// TIA Portal V17 program export: 1 tag tables, 0 data types, 1 data blocks, 1 code blocks (in call order from the OBs), 0 instance data blocks

VAR_GLOBAL   // PLC tag table "红绿灯变量表"
   StartPB AT %M0.0 : Bool;   // HMI 启动按钮
   StopPB AT %M0.1 : Bool;   // HMI 停止按钮
   Run AT %M0.2 : Bool;   // 运行自锁与指示灯
   NS_Red AT %Q0.0 : Bool;   // 南北红灯
   NS_Yellow AT %Q0.1 : Bool;   // 南北黄灯
   NS_Green AT %Q0.2 : Bool;   // 南北绿灯
   EW_Red AT %Q0.3 : Bool;   // 东西红灯
   EW_Yellow AT %Q0.4 : Bool;   // 东西黄灯
   EW_Green AT %Q0.5 : Bool;   // 东西绿灯
   Done1 AT %M1.0 : Bool;   // 东西绿灯定时到
   Done2 AT %M1.1 : Bool;   // 东西黄灯定时到
   Done3 AT %M1.2 : Bool;   // 南北绿灯定时到
   Done4 AT %M1.3 : Bool;   // 南北黄灯定时到
END_VAR

DATA_BLOCK "TrafficTimers"   // DB1
{ S7_Optimized_Access := 'FALSE' }
   VAR
      T1 : TON_TIME;
      T2 : TON_TIME;
      T3 : TON_TIME;
      T4 : TON_TIME;
   END_VAR
BEGIN
END_DATA_BLOCK

ORGANIZATION_BLOCK "Main"   // OB1, LAD, ProgramCycle
{ S7_Optimized_Access := 'TRUE' }
VERSION : 0.1
// stored: AutoNumber true, IsIECCheckEnabled false, SetENOAutomatically false
   VAR_INPUT
      Initial_Call : Bool;   // Initial call of this OB
      Remanence : Bool;   // =True, if remanent data are available
   END_VAR
BEGIN

REGION Network 1: 启停自锁
   // 启动后保持运行，停止优先。
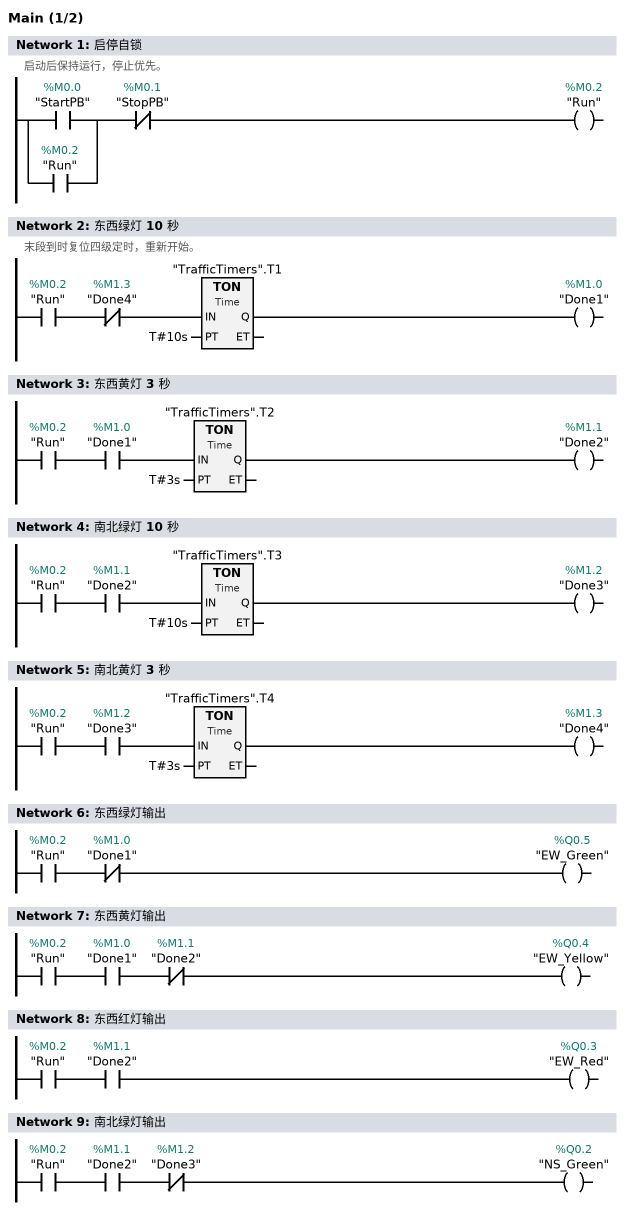
   RUNG wire#powerrail
      Contact( "StartPB" )
      wire#w1
      I_Contact( "StopPB" )
      Coil( "Run" )
   END_RUNG
   RUNG wire#powerrail
      Contact( "Run" )
   END_RUNG wire#w1
   // the same network as SCL:
   "Run" := ("StartPB" OR "Run") AND NOT "StopPB";
END_REGION

REGION Network 2: 东西绿灯 10 秒
   // 末段到时复位四级定时，重新开始。
   RUNG wire#powerrail
      Contact( "Run" )
      I_Contact( "Done4" )
      { S7_Templates := "time_type := Time" } "TrafficTimers".T1.TON(pt := T#10s, et =>)
      Coil( "Done1" )
   END_RUNG
   // the same network as SCL:
   "TrafficTimers".T1.TON(IN := "Run" AND NOT "Done4", PT := T#10s);
   "Done1" := "TrafficTimers".T1.Q;
END_REGION

REGION Network 3: 东西黄灯 3 秒
   RUNG wire#powerrail
      Contact( "Run" )
      Contact( "Done1" )
      { S7_Templates := "time_type := Time" } "TrafficTimers".T2.TON(pt := T#3s, et =>)
      Coil( "Done2" )
   END_RUNG
   // the same network as SCL:
   "TrafficTimers".T2.TON(IN := "Run" AND "Done1", PT := T#3s);
   "Done2" := "TrafficTimers".T2.Q;
END_REGION

REGION Network 4: 南北绿灯 10 秒
   RUNG wire#powerrail
      Contact( "Run" )
      Contact( "Done2" )
      { S7_Templates := "time_type := Time" } "TrafficTimers".T3.TON(pt := T#10s, et =>)
      Coil( "Done3" )
   END_RUNG
   // the same network as SCL:
   "TrafficTimers".T3.TON(IN := "Run" AND "Done2", PT := T#10s);
   "Done3" := "TrafficTimers".T3.Q;
END_REGION

REGION Network 5: 南北黄灯 3 秒
   RUNG wire#powerrail
      Contact( "Run" )
      Contact( "Done3" )
      { S7_Templates := "time_type := Time" } "TrafficTimers".T4.TON(pt := T#3s, et =>)
      Coil( "Done4" )
   END_RUNG
   // the same network as SCL:
   "TrafficTimers".T4.TON(IN := "Run" AND "Done3", PT := T#3s);
   "Done4" := "TrafficTimers".T4.Q;
END_REGION

REGION Network 6: 东西绿灯输出
   RUNG wire#powerrail
      Contact( "Run" )
      I_Contact( "Done1" )
      Coil( "EW_Green" )
   END_RUNG
   // the same network as SCL:
   "EW_Green" := "Run" AND NOT "Done1";
END_REGION

REGION Network 7: 东西黄灯输出
   RUNG wire#powerrail
      Contact( "Run" )
      Contact( "Done1" )
      I_Contact( "Done2" )
      Coil( "EW_Yellow" )
   END_RUNG
   // the same network as SCL:
   "EW_Yellow" := "Run" AND "Done1" AND NOT "Done2";
END_REGION

REGION Network 8: 东西红灯输出
   RUNG wire#powerrail
      Contact( "Run" )
      Contact( "Done2" )
      Coil( "EW_Red" )
   END_RUNG
   // the same network as SCL:
   "EW_Red" := "Run" AND "Done2";
END_REGION

REGION Network 9: 南北绿灯输出
   RUNG wire#powerrail
      Contact( "Run" )
      Contact( "Done2" )
      I_Contact( "Done3" )
      Coil( "NS_Green" )
   END_RUNG
   // the same network as SCL:
   "NS_Green" := "Run" AND "Done2" AND NOT "Done3";
END_REGION

REGION Network 10: 南北黄灯输出
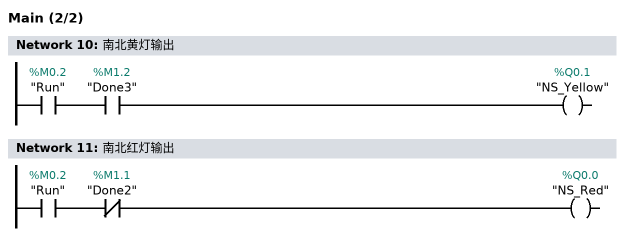
   RUNG wire#powerrail
      Contact( "Run" )
      Contact( "Done3" )
      Coil( "NS_Yellow" )
   END_RUNG
   // the same network as SCL:
   "NS_Yellow" := "Run" AND "Done3";
END_REGION

REGION Network 11: 南北红灯输出
   RUNG wire#powerrail
      Contact( "Run" )
      I_Contact( "Done2" )
      Coil( "NS_Red" )
   END_RUNG
   // the same network as SCL:
   "NS_Red" := "Run" AND NOT "Done2";
END_REGION
END_ORGANIZATION_BLOCK
